Fanuc KAREL source: kt00240.KL

-- PROVISIONAL review KL for V770-1; original PC SHA256 9b4dc21110e25e2cb9fc0c392b7bf8f3ba6ac6bf1a69a320fc60ed74c39b83fe
-- Incomplete behavior may be omitted. Consult companion uncertainty JSON. Do not deploy.
PROGRAM KT00240
%NOLOCKGROUP
VAR
  I1 : INTEGER
  OUT : INTEGER
-- UNRESOLVED_DECL H2 type=002017
BEGIN
  -- UNRESOLVED_PC offsets 5-16; opcodes 2E,23
  -- UNRESOLVED_PC offsets 21-35; opcodes 2E,22,9D,33,B4
  -- UNRESOLVED_PC offsets 40-62; opcodes 21,22,9D,33,B3,47,23
  -- UNRESOLVED_PC offsets 67-71; opcodes 7F
END KT00240
